// TIA Portal V21 export
ORGANIZATION_BLOCK "Pair"   // OB1, LAD
BEGIN

REGION Network 1: Motor
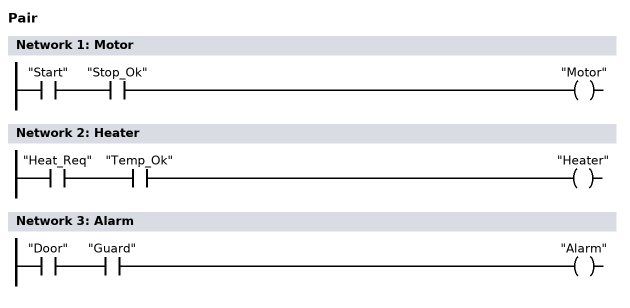
   RUNG wire#powerrail
      Contact( "Start" )
      Contact( "Stop_Ok" )
      Coil( "Motor" )
   END_RUNG
   // the same network as SCL:
   "Motor" := "Start" AND "Stop_Ok";
END_REGION

REGION Network 2: Heater
   RUNG wire#powerrail
      Contact( "Heat_Req" )
      Contact( "Temp_Ok" )
      Coil( "Heater" )
   END_RUNG
   // the same network as SCL:
   "Heater" := "Heat_Req" AND "Temp_Ok";
END_REGION

REGION Network 3: Alarm
   RUNG wire#powerrail
      Contact( "Door" )
      Contact( "Guard" )
      Coil( "Alarm" )
   END_RUNG
   // the same network as SCL:
   "Alarm" := "Door" AND "Guard";
END_REGION
END_ORGANIZATION_BLOCK
